(* IEC 61131-3 sources: repolevel_ST_code_completion/ground_truth/repoeval_traffic_light/readful_result, 4 files *)

(* ---- F_SecondsToTime.st ---- *)
It seems like you are sharing code fragments from a repository related to traffic light control in a PLC programming environment. The code is written in Structured Text (ST), which is commonly used in industrial automation.

The `F_SecondsToTime` function is already defined in the provided code fragments. Here is the complete implementation of the function:

```st
FUNCTION F_SecondsToTime : TIME
VAR_INPUT
	dwSeconds	:	DWORD;		//输入的秒数
END_VAR

// 将秒数（DWORD）转换为TIME类型
// 秒数乘以1000得到毫秒
F_SecondsToTime := DWORD_TO_TIME(dwSeconds * 1000);
```

### Explanation:
- **Purpose**: This function converts a given number of seconds (as a `DWORD`) into a `TIME` data type.
- **Logic**: Since the `TIME` data type in PLC programming typically represents time in milliseconds, the function multiplies the input seconds by 1000 to convert them into milliseconds. It then uses the `DWORD_TO_TIME` conversion function to cast the result into the `TIME` type.

If you have any specific questions or need further assistance with this code or related functionality, feel free to ask!

(* ---- F_SecondsToTime_1.st ---- *)
It seems like you are sharing code fragments from a repository related to traffic light control in a PLC programming environment. The code is written in Structured Text (ST), which is commonly used in industrial automation.

The `F_SecondsToTime` function is already defined in the provided code fragments. Here is the complete implementation of the function:

```st
FUNCTION F_SecondsToTime : TIME
VAR_INPUT
	dwSeconds	:	DWORD;		//输入的秒数
END_VAR

// 将秒数（DWORD）转换为TIME类型
// 秒数乘以1000得到毫秒
F_SecondsToTime := DWORD_TO_TIME(dwSeconds * 1000);
```

### Explanation:
- **Purpose**: This function converts a given number of seconds (as a `DWORD`) into a `TIME` data type.
- **Logic**: Since the `TIME` data type in PLC programming typically represents time in milliseconds, the function multiplies the input seconds by 1000 to convert them into milliseconds. It then uses the `DWORD_TO_TIME` conversion function to cast the result into the `TIME` type.

If you have any specific questions or need further assistance with this code or related functionality, feel free to ask!

(* ---- F_TimeToSeconds.st ---- *)
It seems you are sharing a code snippet for a function `F_TimeToSeconds` and providing context from other files in the repository. Based on the provided information, the function `F_TimeToSeconds` is designed to convert a `TIME` data type (representing a duration in milliseconds) into a `DWORD` (representing the equivalent duration in seconds).

Here is the implementation of the `F_TimeToSeconds` function:

```st
FUNCTION F_TimeToSeconds : DWORD
VAR_INPUT
	tTime	:	TIME;		//输入的时间
END_VAR

// 将TIME类型转换为秒数（DWORD）
// TIME内部是毫秒，除以1000得到秒数
F_TimeToSeconds := DINT_TO_DWORD(TRUNC(TIME_TO_DWORD(tTime) / 1000.0));
```

### Explanation of the Code:
1. **Input Parameter**:
   - `tTime`: A `TIME` type input that represents a duration in milliseconds.

2. **Conversion Logic**:
   - The `TIME_TO_DWORD` function converts the `TIME` value into a `DWORD` representing the duration in milliseconds.
   - Dividing this value by `1000.0` converts the duration from milliseconds to seconds.
   - The `TRUNC` function truncates the result to remove any fractional part, ensuring the result is an integer.
   - The `DINT_TO_DWORD` function converts the truncated integer value into a `DWORD`.

3. **Output**:
   - The function returns the duration in seconds as a `DWORD`.

### Usage in the Repository:
- This function is used in various parts of the repository to convert `TIME` values (e.g., `MGreenTimeOn`, `MGreenTimeFlash`, `MYellowTimeOn`) into seconds for further processing or display. For example:
  - In `TrafficLightHMI`, it is used to initialize variables like `greenTimeOn`, `greenTimeFlash`, and `yellowTimeOn` with the corresponding durations in seconds.

If you have any specific questions or need further clarification, feel free to ask!

(* ---- F_TimeToSeconds_1.st ---- *)
It seems you are sharing a code snippet for a function `F_TimeToSeconds` and providing context from other files in the repository. Based on the provided information, the function `F_TimeToSeconds` is designed to convert a `TIME` data type (representing a duration in milliseconds) into a `DWORD` (representing the equivalent duration in seconds).

Here is the implementation of the `F_TimeToSeconds` function:

```st
FUNCTION F_TimeToSeconds : DWORD
VAR_INPUT
	tTime	:	TIME;		//输入的时间
END_VAR

// 将TIME类型转换为秒数（DWORD）
// TIME内部是毫秒，除以1000得到秒数
F_TimeToSeconds := DINT_TO_DWORD(TRUNC(TIME_TO_DWORD(tTime) / 1000.0));
```

### Explanation of the Code:
1. **Input Parameter**:
   - `tTime`: A `TIME` type input that represents a duration in milliseconds.

2. **Conversion Logic**:
   - The `TIME_TO_DWORD` function converts the `TIME` value into a `DWORD` representing the duration in milliseconds.
   - Dividing this value by `1000.0` converts the duration from milliseconds to seconds.
   - The `TRUNC` function truncates the result to remove any fractional part, ensuring the result is an integer.
   - The `DINT_TO_DWORD` function converts the truncated integer value into a `DWORD`.

3. **Output**:
   - The function returns the duration in seconds as a `DWORD`.

### Usage in the Repository:
- This function is used in various parts of the repository to convert `TIME` values (e.g., `MGreenTimeOn`, `MGreenTimeFlash`, `MYellowTimeOn`) into seconds for further processing or display. For example:
  - In `TrafficLightHMI`, it is used to initialize variables like `greenTimeOn`, `greenTimeFlash`, and `yellowTimeOn` with the corresponding durations in seconds.

If you have any specific questions or need further clarification, feel free to ask!
